TEXTLIST TextList_CIP_Type
  0 = ' '
  1 = 'R Water'
  2 = 'Detergent'
  3 = 'Full'
   = ''
END_TEXTLIST

(* stored: Version 1.1.0.1, ProductVersion 3.1.4024.12
   TextList TextList_CIP_Type: Id {22cd0b7c-8087-48d4-8014-15cbb12b846c} *)
